Yaskawa INFORM job: SPLITTE2.JBI

/JOB
//NAME SPLITTE2
//POS
///NPOS 15,0,0,0,0,0
///TOOL 1
///POSTYPE BASE
///RECTAN
///RCONF 0,0,0,0,0,0,0,0
C00000=674.300,134.999,685.980,-66.22,8.38,-107.67
C00001=661.027,82.386,686.221,-67.04,7.80,-111.79
C00002=674.300,134.999,685.980,-66.22,8.38,-107.67
C00003=661.027,82.386,686.221,-67.04,7.80,-111.79
C00004=674.300,134.999,685.980,-66.22,8.38,-107.67
C00005=661.027,82.386,686.221,-67.04,7.80,-111.79
C00006=674.300,134.999,685.980,-66.22,8.38,-107.67
C00007=661.027,82.386,686.221,-67.04,7.80,-111.79
C00008=674.300,134.999,685.980,-66.22,8.38,-107.67
C00009=661.027,82.386,686.221,-67.04,7.80,-111.79
C00010=674.300,134.999,685.980,-66.22,8.38,-107.67
C00011=661.027,82.386,686.221,-67.04,7.80,-111.79
C00012=674.300,134.999,685.980,-66.22,8.38,-107.67
C00013=661.027,82.386,686.221,-67.04,7.80,-111.79
C00014=674.300,134.999,685.980,-66.22,8.38,-107.67
//INST
///DATE 2026/10/26 01:19
///COMM Generated using RoboDK
///ATTR SC,RW,RJ
///GROUP1 RB1
NOP
MOVL C00000 V=200.0
MOVL C00001 V=200.0
MOVL C00002 V=200.0
MOVL C00003 V=200.0
MOVL C00004 V=200.0
MOVL C00005 V=200.0
MOVL C00006 V=200.0
MOVL C00007 V=200.0
MOVL C00008 V=200.0
MOVL C00009 V=200.0
MOVL C00010 V=200.0
MOVL C00011 V=200.0
MOVL C00012 V=200.0
MOVL C00013 V=200.0
MOVL C00014 V=200.0
END
